# B&R Automation Studio project Starter
Automation Studio 4.12.1; Virtual PLC training example; no physical controller connection

## Configuration Example

### Task classes (CPU.sw)
```
Cyclic#1 (cycle 10000 us):
  Main <- Main.prg
```

### Hardware
```
CPU : VirtualTrainingCPU
  Cyclic1Duration = 10000
```

## Logical view

### Global.var
```iecst
VAR_GLOBAL
    StartCommand : BOOL := FALSE;
    StopCommand : BOOL := FALSE;
    DoorClosed : BOOL := TRUE;
    ResetCounter : BOOL := FALSE;
    MotorRunning : BOOL := FALSE;
    ScanCounter : DINT := 0;
END_VAR
```

### Program Logical/Main (IEC)

#### MainCyclic.st
```iecst
PROGRAM _CYCLIC
(* Training logic only. Commands and outputs share the virtual memory. *)
MotorRunning := StartCommand AND NOT StopCommand AND DoorClosed;
IF ResetCounter THEN
    ScanCounter := 0;
ELSIF MotorRunning THEN
    ScanCounter := ScanCounter + 1;
END_IF;
END_PROGRAM
```
